Fanuc KAREL source: KT00890.KL

PROGRAM KT00890
%NOLOCKGROUP
VAR
  P1: XYZWPREXT
  P2: XYZWPREXT
  OUT: POSITION
BEGIN
  P1.X = 1.0
  P2.Y = 2.0
  P1.X = 1.0
  P2.Y = 2.0
  OUT = INV(P1)
END KT00890
